Fanuc TP program (LS listing): MainCa.LS

/PROG  MainCa
/ATTR
OWNER		= MNEDITOR;
COMMENT		= "RoboDK sequence";
PROG_SIZE	= 0;
CREATE		= DATE 31-12-14  TIME 12:00:00;
MODIFIED	= DATE 31-12-14  TIME 12:00:00;
FILE_NAME	= MainCa;
VERSION		= 0;
LINE_COUNT	= 14;
MEMORY_SIZE	= 0;
PROTECT		= READ_WRITE;
TCD:  STACK_SIZE	= 0,
      TASK_PRIORITY	= 50,
      TIME_SLICE	= 0,
      BUSY_LAMP_OFF	= 0,
      ABORT_REQUEST	= 0,
      PAUSE_REQUEST	= 0;
DEFAULT_GROUP	= 1,*,*,*,*;
CONTROL_CODE	= 00000000 00000000;
/MN
   1:  ! Program generated by RoboDK v6.0.7 for Fanuc M-1iA/0.5S on XX ;
   2:  ! /XX/XXXX 18:00:00 ;
   3:  ! Using nominal kinematics. ;
   4:  PR[9,1]=1234.570 ;
   5:  PR[9,2]=-98.765 ;
   6:  PR[9,3]=50.500 ;
   7:  PR[9,4]=0.000 ;
   8:  PR[9,5]=0.000 ;
   9:  PR[9,6]=30.000 ;
  10:  UFRAME[9]=PR[9] ;
  11:  UFRAME_NUM=9 ;
  12:J P[1] 20% FINE ;
  13:  CALL SubProg2 ;
  14:  CALL NotAProg ;
/POS
P[1]{
   GP1:
    UF : 9, UT : 9,
	J1=    10.000000 deg,	J2=    -20.000000 deg,	J3=    50.000000  mm,
	J4=    30.000000 deg
};
/END
